Fanuc KAREL source: KT00806.KL

PROGRAM KT00806
%NOLOCKGROUP
VAR
  S1: STRING[80]
  S2: STRING[80]
  OUT: INTEGER
BEGIN
  S1 = 'A'
  S2 = 'B'
  S1 = 'A'
  S2 = 'B'
  OUT = EXP(S1)
END KT00806
